{region 'Documentation'}
(*!
<summary>Check that the token count is outside the inclusive Minimum..Maximum range.</summary>
<description>

StartIndex is an absolute declared IN index, not an offset. Length selects 1..255
elements; the complete selected range must fit IN. Invalid references or ranges report
Error.

Keep supplied arrays stable for the call. Input data is read, not copied or retained as a
snapshot.

Comparison applies Mask to both values; bits outside it are ignored. The default mask
selects all bits.

Counts the currently selected region on evaluation, not occurrences across cycles.
TokenCount exposes the last computed count. Inclusive range bounds must be ordered; reversed
bounds report Error.

The value token matches under Mask; bits outside Mask are ignored.

</description>
*)
{endregion}
FUNCTION_BLOCK AssertValueTokenCntNotInRange_Word EXTENDS AssertionBase
VAR_INPUT
    StartIndex : DINT; //! First selected index in IN; uses the array's declared index range, not a zero-based offset.
    Length : USINT; //! Number of selected elements starting at StartIndex; must fit the array range; valid range 1..255.
    Minimum : UINT; //! Inclusive lower bound of the comparison; for a range, must not exceed Maximum.
    Maximum : UINT; //! Inclusive upper bound of the comparison; for a range, must not be below Minimum.
    Token : WORD; //! Value searched for in the selected range; Mask selects the compared bits.
    Mask : WORD := WORD#16#FFFF; //! Bits included in the comparison; bits outside the mask are ignored.
END_VAR
VAR_IN_OUT CONSTANT
    IN : ARRAY[*] OF WORD; //! Keep the searched data stable during the call.
END_VAR
VAR
    FTokenCount : UINT;
END_VAR

SUPER^();

{region 'Documentation'}
(*!
<summary>Validate configuration, count tokens and apply the count predicate.</summary>
*)
{endregion}
METHOD PROTECTED Assert
VAR
    InLowerIndex : DINT;
    InUpperIndex : DINT;
    EndIndex : LINT;
    Message : STRING(GVL_Constants.MessageLength);
END_VAR
VAR CONSTANT
    HexDigitCount : USINT := 4;
END_VAR
IF NOT EvaluationActive THEN
    RETURN;
END_IF;

IF Result = E_Result.Error THEN
    RETURN;
END_IF;

// C0371: FB input is checked before any reference access.
{warning disable C0371}
IF NOT __ISVALIDREF(IN) THEN
    FTokenCount := 0;
    Error(Message := 'Assertion error: IN reference is invalid.');
    RETURN;
END_IF;

InLowerIndex := LOWER_BOUND(IN, 1);
InUpperIndex := UPPER_BOUND(IN, 1);
EndIndex := DINT_TO_LINT(StartIndex) + USINT_TO_LINT(Length) - 1;
IF (Length = 0)
    OR (StartIndex < InLowerIndex) OR (StartIndex > InUpperIndex)
    OR (EndIndex > DINT_TO_LINT(InUpperIndex)) THEN
    FTokenCount := 0;
    Message := CONCAT('Assertion error: invalid search range. StartIndex = ',
        DINT_TO_STRING(StartIndex));
    Message := CONCAT(Message, ', Length = ');
    Message := CONCAT(Message, USINT_TO_STRING(Length));
    Error(Message := Message);
    RETURN;
END_IF;

IF Minimum > Maximum THEN
    FTokenCount := 0;
    Message := CONCAT('Assertion error: reversed token count bounds. Minimum = ',
        UINT_TO_STRING(Minimum));
    Message := CONCAT(Message, ', Maximum = ');
    Message := CONCAT(Message, UINT_TO_STRING(Maximum));
    Error(Message := Message);
    RETURN;
END_IF;

IF Result = E_Result.Failed THEN
    RETURN;
END_IF;

FTokenCount := CountValueTokens_Word(StartIndex := StartIndex,
    Length := Length,
    Token := Token,
    Mask := Mask,
    IN := IN);

IF (FTokenCount >= Minimum) AND (FTokenCount <= Maximum) THEN
    Message := CONCAT('Assertion failed: value token count violates NotInRange. Actual = ',
        UINT_TO_STRING(FTokenCount));
    Message := CONCAT(Message, ', Minimum = ');
    Message := CONCAT(Message, UINT_TO_STRING(Minimum));
    Message := CONCAT(Message, ', Maximum = ');
    Message := CONCAT(Message, UINT_TO_STRING(Maximum));
    Message := CONCAT(Message, ', Token = ');
    Message := CONCAT(Message, CreateAssertionTextValue_Hex(Value := WORD_TO_LWORD(Token),
        DigitCount := HexDigitCount));
    Message := CONCAT(Message, ', Mask = ');
    Message := CONCAT(Message, CreateAssertionTextValue_Hex(Value := WORD_TO_LWORD(Mask),
        DigitCount := HexDigitCount));
    Fail(Message := Message);
    RETURN;
END_IF;

Pass();
{warning restore C0371}
END_METHOD

{region 'Documentation'}
(*!
<summary>Clear the retained count on framework reset.</summary>
*)
{endregion}
METHOD PROTECTED ResetAssertion
FTokenCount := 0;
END_METHOD

{region 'Documentation'}
(*!
<summary>Return the most recently evaluated token count.</summary>
<description>

Counts occurrences in one selected array region, not across PLC cycles. Retained while
disabled or after Failed; reset and detected configuration errors clear it. Reading this
property does not search the array.

</description>
*)
{endregion}
{attribute 'monitoring' := 'call'}
PROPERTY PUBLIC TokenCount : UINT //! Return the most recently evaluated token count.
GET // PUBLIC
TokenCount := FTokenCount;
END_GET
END_PROPERTY

END_FUNCTION_BLOCK

(* stored: Version 1.1.0.1
   POU AssertValueTokenCntNotInRange_Word: Id {cd7cb081-2b08-42a4-8768-ab249f810170}, SpecialFunc None
   Folder Internal: Id {3cc2702f-908c-4e55-af72-7920c05b04d6}
   Method Assert: Id {85f1b081-b5bf-4d6f-a6d4-2452d156e9d7}
   Method ResetAssertion: Id {b900c246-2b0c-4a60-b1d3-d7891c7913ff}
   Property TokenCount: Id {f2dabcf4-a167-403a-821e-b824b91fa057}
   Get Get: Id {9f1a8775-a179-4d96-81af-ad0d256fb314} *)
